// TIA Portal V20 export
VAR_GLOBAL   // PLC tag table "PLC-A3-DQ"
   "-KA1" AT %Q0.0 : Bool;   // OSVĚTLENÍ FOLIE
   "-KA2" AT %Q0.1 : Bool;   // OSVĚTLENÍ FOLIE
   "-KA3" AT %Q0.2 : Bool;   // OSVĚTLENÍ FOLIE
   "-KA4" AT %Q0.3 : Bool;   // OSVĚTLENÍ ETIKETA
   "-KA5" AT %Q0.4 : Bool;   // OSVĚTLENÍ ETIKETA
   "-KA18" AT %Q0.5 : Bool;   // MAJÁK_žlutá
   "-KA19" AT %Q0.6 : Bool;   // MAJÁK_červená
   "-KA20" AT %Q0.7 : Bool;   // MAJÁK_zelena
   "-KA21" AT %Q1.0 : Bool;   // HOUKAČKA
   RESERVE_DQ AT %Q1.1 : Bool;
END_VAR
